Staubli VAL3: io.dtx

mdesc mNomSpeed
public dio dInput[64]
public dio dOutput[64]
public aio aInput[16]
public aio aOutput[16]
